(* IEC 61131-3 sources: daoli-st-library/_quarantine/R79, 13 files *)

(* ---- FC_DL_CalIsLeapYear.st ---- *)
(*==============================================================================
 * 组件名称 : FC_DL_CalIsLeapYear ｜ 子库 : DL_MathData ｜ v1.0.0 ｜ 2026-11-24
 * 平台     : CODESYS 3.5 / TwinCAT 3 / InoProShop / Machine Expert（纯 IEC，无厂商库）
 * 功能简介 : 公历（格里高利历）闰年判定 —— 能被 4 整除且不能被 100 整除，或能被 400
 *            整除即为闰年。纯整数取余，无浮点、无日历库依赖。
 * 契约     : 返回 TRUE=闰年；nYear < 1583（格里高利历起点）返回 FALSE 且
 *            bValid := FALSE —— 儒略历闰年口径与本件不同，域外一律不认。
 *            纯函数无状态，同输入同输出。
 * 依赖     : 无 DL_ 内部依赖（R16 自足实现），无标准库函数调用
 * 错误码   : R297 零码位范式：eErr 恒 0，仅以 bError / bValid 表达（本件结构性不置 bError）
 * 红线自检 : R1 零全局 R2 零%I/%Q R3 纯IEC R4 取余无除法歧义、域闸先判年份
 *            R5 双语注释 R6 N/A（无状态机）R7 N/A（无定时器/沿实例）
 *            R10 无类型转换 R11 全声明行分号 R15 标识符零保留字冲突 R18 N/A（无 bReset）
 * 修订历史 : 2026-11-24 R79-A 首版（日历算术族 1/9）
 *============================================================================*)
FUNCTION FC_DL_CalIsLeapYear : BOOL
VAR_INPUT
    nYear    : DINT;    // 待判定公历年，有效域 1583 及以上 [年] / Gregorian year to test, valid from 1583 [year]
END_VAR
VAR_OUTPUT
    eErr     : UDINT;   // 错误码，零码位范式恒 0 / error id, always zero under the zero-code rule
    bError   : BOOL;    // 故障标志，本件结构性不置位 / fault flag, never raised by this component
    bValid   : BOOL;    // 年份落在格里高利历域内为真 / TRUE when the year is inside the Gregorian domain
END_VAR
VAR CONSTANT
    DL_GREG_START : DINT := 1583;   // 格里高利历起点年 [年] / first Gregorian year [year]
    DL_STEP4      : DINT := 4;      // 闰年基本步长 [年] / base leap step [year]
    DL_STEP100    : DINT := 100;    // 世纪基数 [年] / century radix [year]
    DL_STEP400    : DINT := 400;    // 四世纪基数 [年] / four century radix [year]
    DL_ZERO       : DINT := 0;      // 整数零哨兵 [无量纲] / integer zero sentinel [dimensionless]
END_VAR
VAR
    nMod4    : DINT;    // 年份除 4 的余数 [无量纲] / remainder of the year divided by four [dimensionless]
    nMod100  : DINT;    // 年份除 100 的余数 [无量纲] / remainder of the year divided by one hundred [dimensionless]
    nMod400  : DINT;    // 年份除 400 的余数 [无量纲] / remainder of the year divided by four hundred [dimensionless]
END_VAR

// 段 1｜出口预置：任何路径下结果确定 / segment 1, preset the exit so that every path is deterministic
FC_DL_CalIsLeapYear := FALSE;   // 缺省非闰年 / default is not a leap year
eErr   := 0;                    // 零码位范式 / zero-code rule
bError := FALSE;                // 本件不产生故障级 / this component raises no fault
bValid := FALSE;                // 域闸通过前不认结果 / the result stays unusable until the domain gate passes

// 段 2｜域闸：1583 之前属儒略历，闰年口径不同，直接拒绝 / segment 2, the domain gate rejects years before 1583
IF nYear < DL_GREG_START THEN
    RETURN;                     // 返回 FALSE 且 bValid 保持 FALSE / return FALSE with bValid still FALSE
END_IF
bValid := TRUE;                 // 年份入域，结果可用 / the year is inside the domain, the result is usable

// 段 3｜闰年判据：先取三个余数，再做布尔合成（避免重复取余） / segment 3, the leap rule on three remainders
nMod4   := nYear MOD DL_STEP4;      // 4 年周期余数 / remainder against four years
nMod100 := nYear MOD DL_STEP100;    // 100 年周期余数 / remainder against one hundred years
nMod400 := nYear MOD DL_STEP400;    // 400 年周期余数 / remainder against four hundred years
IF ((nMod4 = DL_ZERO) AND (nMod100 <> DL_ZERO)) OR (nMod400 = DL_ZERO) THEN
    FC_DL_CalIsLeapYear := TRUE;    // 整除 4 且不整除 100，或整除 400 / divisible by four but not by one hundred, or divisible by four hundred
END_IF
END_FUNCTION

(* ---- FC_DL_CalIsoWeekNo.st ---- *)
(*==============================================================================
 * 组件名称 : FC_DL_CalIsoWeekNo ｜ 子库 : DL_MathData ｜ v1.0.0 ｜ 2026-11-24
 * 平台     : CODESYS 3.5 / TwinCAT 3 / InoProShop / Machine Expert（纯 IEC，无厂商库）
 * 功能简介 : ISO 8601 周号 —— 周一起算，含 1 月 4 日的那一周为第 1 周。核心式
 *            week = (年内序号 − ISO 星期 + 10) DIV 7。跨年归属单独处理：算出 0 即属
 *            上年末周，算出超过当年周数即属次年 W1，并用出参 nWeekYear 标明归属年。
 * 契约     : 返回周号 1~53，nWeekYear 为归属年；nYear < 1583、月份或日越界时返回 -1、
 *            bError := TRUE、nWeekYear := 0。纯函数无状态。
 * 依赖     : 无 DL_ 内部依赖（R16 自足实现），无标准库函数调用
 * 错误码   : R297 零码位范式：eErr 恒 0，仅以 bError / bValid 表达
 * 红线自检 : R1 零全局 R2 零%I/%Q R3 纯IEC R4 三层域闸、取余操作数恒非负、除数为常量 7
 *            R5 双语注释 R6 N/A（无状态机）R7 N/A（无定时器/沿实例）
 *            R10 无类型转换 R11 全声明行分号 R15 标识符零保留字冲突 R18 N/A（无 bReset）
 * 遗留假设 : 53 周年判据按 ISO 官方口径取「1 月 1 日为周四」或「闰年且 1 月 1 日为周三」；
 *            该两式与「12 月 31 日落在第 53 周」等价，本件用前者以便直接复用 1 月 1 日序数。
 * 修订历史 : 2026-11-24 R79-A 首版（日历算术族 6/9）
 *============================================================================*)
FUNCTION FC_DL_CalIsoWeekNo : DINT
VAR_INPUT
    nYear      : DINT;  // 公历年，域闸 1583 及以上 [年] / Gregorian year, domain starts at 1583 [year]
    nMonth     : DINT;  // 月份 1~12 [月] / month from one to twelve [month]
    nDay       : DINT;  // 日 1~当月天数 [天] / day from one to the month length [day]
END_VAR
VAR_OUTPUT
    eErr       : UDINT; // 错误码，零码位范式恒 0 / error id, always zero under the zero-code rule
    bError     : BOOL;  // 日期非法或域外为真 / TRUE when the date is illegal or out of domain
    bValid     : BOOL;  // 结果可用标志 / result usable flag
    nWeekYear  : DINT;  // 周号归属年，故障时 0 [年] / year owning the ISO week, zero on fault [year]
END_VAR
VAR CONSTANT
    DL_GREG_START : DINT := 1583;   // 格里高利历起点年 [年] / first Gregorian year [year]
    DL_MONTH_MIN  : DINT := 1;      // 月份与日的下界 [月] / lower bound of the month and the day [month]
    DL_MONTH_MAX  : DINT := 12;     // 月份上界 [月] / upper month bound [month]
    DL_DAYS_COMMON : DINT := 365;   // 平年天数 [天] / days in a common year [day]
    DL_DAYS_FEB   : DINT := 28;     // 平年 2 月天数 [天] / February days in a common year [day]
    DL_DAYS_30    : DINT := 30;     // 小月天数 [天] / days in a short month [day]
    DL_DAYS_31    : DINT := 31;     // 大月天数 [天] / days in a long month [day]
    DL_STEP4      : DINT := 4;      // 闰年基本步长 [年] / base leap step [year]
    DL_STEP100    : DINT := 100;    // 世纪基数 [年] / century radix [year]
    DL_STEP400    : DINT := 400;    // 四世纪基数 [年] / four century radix [year]
    DL_WEEK_MOD   : DINT := 7;      // 星期与周号的基数 [天] / weekday and week radix [day]
    DL_WEEK_MIN   : DINT := 1;      // 周号下界 [周] / lower bound of the week number [week]
    DL_WEEK_BASE  : DINT := 52;     // 每年基础周数，53 周为特例 [周] / base weeks per year, fifty three is the exception [week]
    DL_WEEK_OFF   : DINT := 10;     // 周号式的固定偏移 [天] / fixed offset of the week formula [day]
    DL_JAN1_DOW53A : DINT := 4;     // 1 月 1 日周四 → 53 周 [星期序号] / Thursday first of January gives fifty three weeks
    DL_JAN1_DOW53B : DINT := 3;     // 闰年 1 月 1 日周三 → 53 周 [星期序号] / Wednesday first of January in a leap year gives fifty three weeks
    DL_ZERO       : DINT := 0;      // 整数零哨兵 [无量纲] / integer zero sentinel [dimensionless]
END_VAR
VAR
    bLeap      : BOOL;  // 当年是否闰年 / whether the year is a leap year
    bLeapPrev  : BOOL;  // 上一年是否闰年 / whether the previous year is a leap year
    nDaysInMon : DINT;  // 当月实际天数 [天] / actual length of the month [day]
    nDaysYear  : DINT;  // 当年总天数 365 或 366 [天] / total days of the year [day]
    nDaysPrev  : DINT;  // 上年总天数 365 或 366 [天] / total days of the previous year [day]
    nA         : DINT;  // 月份压缩偏置 0 或 1 / month compression offset, zero or one
    nY2        : DINT;  // 儒略式内的世纪内年份 / shifted year inside the Julian formula
    nM2        : DINT;  // 儒略式内的三月基月份 / March based month inside the Julian formula
    nJdn       : DINT;  // 目标日期的儒略日序数 [日] / Julian day number of the requested date [day]
    nJdnJan1   : DINT;  // 同年 1 月 1 日的儒略日序数 [日] / Julian day number of January the first [day]
    nDowJan1   : DINT;  // 1 月 1 日的 ISO 星期 1~7 [星期序号] / ISO weekday of January the first, one to seven
    nW         : DINT;  // 目标日期的 ISO 星期 1~7 [星期序号] / ISO weekday of the requested date, one to seven
    nOrd       : DINT;  // 年内序号 1~366 [天] / day of year, one to three hundred sixty six [day]
    nWeek      : DINT;  // 周号中间量 0~54 [周] / week interim value, zero to fifty four [week]
    nWeeksYear : DINT;  // 当年 ISO 周数 52 或 53 [周] / ISO weeks in the year, fifty two or fifty three [week]
END_VAR

// 段 1｜出口预置 / segment 1, preset the exit
FC_DL_CalIsoWeekNo := -1;       // 缺省无效哨兵 / default invalid sentinel
eErr       := 0;                // 零码位范式 / zero-code rule
bError     := FALSE;            // 预置无故障 / preset no fault
bValid     := FALSE;            // 域闸前不认结果 / unusable until the domain gates pass
nWeekYear  := 0;                // 归属年清零 / clear the owning year

// 段 2｜域闸：年份 → 月份 → 日（含闰年 2 月） / segment 2, the three domain gates
bLeap := (((nYear MOD DL_STEP4) = DL_ZERO) AND ((nYear MOD DL_STEP100) <> DL_ZERO)) OR ((nYear MOD DL_STEP400) = DL_ZERO);
nDaysYear := DL_DAYS_COMMON;
IF bLeap THEN
    nDaysYear := DL_DAYS_COMMON + 1;    // 闰年多一天 / a leap year carries one extra day
END_IF
IF (nYear < DL_GREG_START) OR (nMonth < DL_MONTH_MIN) OR (nMonth > DL_MONTH_MAX) THEN
    bError := TRUE;             // 年份或月份越界 / the year or the month is out of range
    RETURN;
END_IF
IF nMonth = 2 THEN
    nDaysInMon := DL_DAYS_FEB;          // 平年 2 月 / common February
    IF bLeap THEN
        nDaysInMon := DL_DAYS_FEB + 1;  // 闰年 2 月 / leap February
    END_IF
ELSIF (nMonth = 4) OR (nMonth = 6) OR (nMonth = 9) OR (nMonth = 11) THEN
    nDaysInMon := DL_DAYS_30;           // 小月 / short month
ELSE
    nDaysInMon := DL_DAYS_31;           // 大月 / long month
END_IF
IF (nDay < DL_MONTH_MIN) OR (nDay > nDaysInMon) THEN
    bError := TRUE;             // 日超出当月天数 / the day exceeds the month length
    RETURN;
END_IF

// 段 3｜两个儒略日序数：目标日期与同年 1 月 1 日 / segment 3, two Julian day numbers
nA   := (14 - nMonth) / 12;                                  // 1、2 月折入上一年 / January and February fold backwards
nY2  := nYear + 4800 - nA;                                   // 世纪内年份偏置 / shifted year
nM2  := nMonth + 12 * nA - 3;                                // 三月基月份 / March based month
nJdn := nDay + (153 * nM2 + 2) / 5 + 365 * nY2 + nY2 / DL_STEP4 - nY2 / DL_STEP100 + nY2 / DL_STEP400 - 32045;
nJdnJan1 := 307 + 365 * (nYear + 4799) + (nYear + 4799) / DL_STEP4 - (nYear + 4799) / DL_STEP100 + (nYear + 4799) / DL_STEP400 - 32045;
nOrd := nJdn - nJdnJan1 + 1;                                 // 年内序号 / day of year
nW   := (nJdn MOD DL_WEEK_MOD) + 1;                           // ISO 星期 1=周一 … 7=周日 / ISO weekday

// 段 4｜周号主式与当年周数：53 周须 1 月 1 日为周四，或闰年且为周三 / segment 4, the week formula and the year length
nWeek := (nOrd - nW + DL_WEEK_OFF) / DL_WEEK_MOD;             // 0~54 中间值 / interim value
nDowJan1 := (nJdnJan1 MOD DL_WEEK_MOD) + 1;                   // 1 月 1 日的 ISO 星期 / ISO weekday of January the first
nWeeksYear := DL_WEEK_BASE;                                   // 缺省 52 周 / default fifty two weeks
IF (nDowJan1 = DL_JAN1_DOW53A) OR (bLeap AND (nDowJan1 = DL_JAN1_DOW53B)) THEN
    nWeeksYear := DL_WEEK_BASE + 1;                           // 该年为 53 周 / the year carries fifty three weeks
END_IF

// 段 5｜跨年归属：0 归上年末周，超年周数归次年 W1 / segment 5, the two cross year branches
nWeekYear := nYear;
IF nWeek < DL_WEEK_MIN THEN
    bLeapPrev := ((((nYear - 1) MOD DL_STEP4) = DL_ZERO) AND (((nYear - 1) MOD DL_STEP100) <> DL_ZERO)) OR (((nYear - 1) MOD DL_STEP400) = DL_ZERO);
    nDaysPrev := DL_DAYS_COMMON;
    IF bLeapPrev THEN
        nDaysPrev := DL_DAYS_COMMON + 1;    // 上年为闰年 / the previous year is a leap year
    END_IF
    nWeek     := (nOrd + nDaysPrev - nW + DL_WEEK_OFF) / DL_WEEK_MOD;   // 换算到上年的序数 / rebase onto the previous year
    nWeekYear := nYear - 1;                                             // 归属上年 / owned by the previous year
ELSIF nWeek > nWeeksYear THEN
    nWeek     := (nOrd - nDaysYear - nW + DL_WEEK_OFF) / DL_WEEK_MOD;   // 换算到次年的序数 / rebase onto the next year
    IF nWeek < DL_WEEK_MIN THEN
        nWeek := DL_WEEK_MIN;                                          // 结构性必为 1，兜底防御 / always one, kept as a guard
    END_IF
    nWeekYear := nYear + 1;                                             // 归属次年 / owned by the next year
END_IF

// 段 6｜出口 / segment 6, exit
FC_DL_CalIsoWeekNo := nWeek;    // 1~53 / one to fifty three
bValid := TRUE;                 // 结果可用 / the result is usable
END_FUNCTION

(* ---- FC_DL_CalMonthDays.st ---- *)
(*==============================================================================
 * 组件名称 : FC_DL_CalMonthDays ｜ 子库 : DL_MathData ｜ v1.0.0 ｜ 2026-11-24
 * 平台     : CODESYS 3.5 / TwinCAT 3 / InoProShop / Machine Expert（纯 IEC，无厂商库）
 * 功能简介 : 给定公历年月，返回该月天数；2 月按闰年判据取 28 或 29，其余月固定 30/31。
 *            纯整数实现，闰年判据内联自足，不调用同族其他件。
 * 契约     : 返回 1~31 为合法天数；nMonth 越界（<1 或 >12）返回 0 且 bError := TRUE。
 *            nYear < 1583 时 2 月按非闰年（28）计数 —— 儒略历口径不入本件，见遗留假设。
 * 依赖     : 无 DL_ 内部依赖（R16 自足实现），无标准库函数调用
 * 错误码   : R297 零码位范式：eErr 恒 0，仅以 bError / bValid 表达
 * 红线自检 : R1 零全局 R2 零%I/%Q R3 纯IEC R4 月份域闸先行、取余无除零面
 *            R5 双语注释 R6 N/A（无状态机）R7 N/A（无定时器/沿实例）
 *            R10 无类型转换 R11 全声明行分号 R15 标识符零保留字冲突 R18 N/A（无 bReset）
 * 遗留假设 : 格里高利历起点之前的 2 月按 28 天计；该域需 29 天的场合请先自查历法归属。
 * 修订历史 : 2026-11-24 R79-A 首版（日历算术族 2/9）
 *============================================================================*)
FUNCTION FC_DL_CalMonthDays : DINT
VAR_INPUT
    nYear     : DINT;   // 公历年，仅供 2 月闰年判定 [年] / Gregorian year used by the February leap test [year]
    nMonth    : DINT;   // 月份 1~12，越界即故障 [月] / month from one to twelve, out of range is a fault [month]
END_VAR
VAR_OUTPUT
    eErr      : UDINT;  // 错误码，零码位范式恒 0 / error id, always zero under the zero-code rule
    bError    : BOOL;   // 月份越界为真，返回 0 / TRUE when the month is out of range, the result is zero
    bValid    : BOOL;   // 结果可用标志 / result usable flag
END_VAR
VAR CONSTANT
    DL_MONTH_MIN  : DINT := 1;      // 月份下界 [月] / lower month bound [month]
    DL_MONTH_MAX  : DINT := 12;     // 月份上界 [月] / upper month bound [month]
    DL_DAYS_31    : DINT := 31;     // 大月天数 [天] / days in a long month [day]
    DL_DAYS_30    : DINT := 30;     // 小月天数 [天] / days in a short month [day]
    DL_DAYS_FEB   : DINT := 28;     // 平年 2 月天数 [天] / February days in a common year [day]
    DL_GREG_START : DINT := 1583;   // 格里高利历起点年 [年] / first Gregorian year [year]
    DL_STEP4      : DINT := 4;      // 闰年基本步长 [年] / base leap step [year]
    DL_STEP100    : DINT := 100;    // 世纪基数 [年] / century radix [year]
    DL_STEP400    : DINT := 400;    // 四世纪基数 [年] / four century radix [year]
    DL_ZERO       : DINT := 0;      // 整数零哨兵 [无量纲] / integer zero sentinel [dimensionless]
END_VAR
VAR
    bLeap     : BOOL;   // 当年是否闰年 / whether the year is a leap year
END_VAR

// 段 1｜出口预置 / segment 1, preset the exit
FC_DL_CalMonthDays := 0;        // 缺省 0 天 / default zero days
eErr   := 0;                    // 零码位范式 / zero-code rule
bError := FALSE;                // 预置无故障 / preset no fault
bValid := FALSE;                // 域闸前不认结果 / unusable until the domain gate passes

// 段 2｜月份域闸：唯一故障出口 / segment 2, the month domain gate is the only fault exit
IF (nMonth < DL_MONTH_MIN) OR (nMonth > DL_MONTH_MAX) THEN
    bError := TRUE;             // 月份越界 / the month is out of range
    RETURN;                     // 返回 0 / return zero
END_IF
bValid := TRUE;                 // 月份入域 / the month is inside the domain

// 段 3｜闰年判据（内联自足，不跨件调用） / segment 3, the leap test implemented inline
bLeap := FALSE;
IF nYear >= DL_GREG_START THEN
    bLeap := (((nYear MOD DL_STEP4) = DL_ZERO) AND ((nYear MOD DL_STEP100) <> DL_ZERO)) OR ((nYear MOD DL_STEP400) = DL_ZERO);
END_IF

// 段 4｜月长选择：2 月单列，30 天月枚举，其余一律 31 天 / segment 4, month length selection
IF nMonth = 2 THEN
    IF bLeap THEN
        FC_DL_CalMonthDays := DL_DAYS_FEB + 1;     // 闰年 2 月 29 天 / twenty nine days in a leap February
    ELSE
        FC_DL_CalMonthDays := DL_DAYS_FEB;         // 平年 2 月 28 天 / twenty eight days otherwise
    END_IF
ELSIF (nMonth = 4) OR (nMonth = 6) OR (nMonth = 9) OR (nMonth = 11) THEN
    FC_DL_CalMonthDays := DL_DAYS_30;              // 4/6/9/11 月为 30 天 / thirty day months
ELSE
    FC_DL_CalMonthDays := DL_DAYS_31;              // 其余为 31 天 / the rest have thirty one days
END_IF
END_FUNCTION

(* ---- FC_DL_CalMonthEndDate.st ---- *)
(*==============================================================================
 * 组件名称 : FC_DL_CalMonthEndDate ｜ 子库 : DL_MathData ｜ v1.0.1 ｜ 2026-11-24
 * 平台     : CODESYS 3.5 / TwinCAT 3 / InoProShop / Machine Expert（纯 IEC，无厂商库）
 * 功能简介 : 给定公历年月，出参返回该月最后一天的日号（月末日期）。月度报表切日、
 *            月累计清零、月末结账触发都以本件为唯一口径。2 月按闰年判据取 28 / 29。
 * 契约     : 合法时返回 TRUE 并写出 nLastDay（1~31）；nMonth 越界或 nYear < 1583 时
 *            返回 FALSE、bError := TRUE、nLastDay := 0。纯函数无状态。
 * 依赖     : 无 DL_ 内部依赖（R16 自足实现），无标准库函数调用
 * 错误码   : R297 零码位范式：eErr 恒 0，仅以 bError / bValid 表达
 * 红线自检 : R1 零全局 R2 零%I/%Q R3 纯IEC R4 年份与月份双域闸、取余无除零面
 *            R5 双语注释 R6 N/A（无状态机）R7 N/A（无定时器/沿实例）
 *            R10 无类型转换 R11 全声明行分号 R15 标识符零保留字冲突 R18 N/A（无 bReset）
 * 修订历史 : 2026-11-24 R79-A 首版（日历算术族 9/9）
 *            2026-11-24  v1.0.1  R79/P4：补年份上界闸 DL_GREG_LAST=9999（原仅下界 1583）
 *============================================================================*)
FUNCTION FC_DL_CalMonthEndDate : BOOL
VAR_INPUT
    nYear     : DINT;   // 公历年，域闸 1583 及以上 [年] / Gregorian year, domain starts at 1583 [year]
    nMonth    : DINT;   // 月份 1~12 [月] / month from one to twelve [month]
END_VAR
VAR_OUTPUT
    eErr      : UDINT;  // 错误码，零码位范式恒 0 / error id, always zero under the zero-code rule
    bError    : BOOL;   // 年份或月份越界为真 / TRUE when the year or the month is out of range
    bValid    : BOOL;   // 出参可用标志 / TRUE when the output is usable
    nLastDay  : DINT;   // 该月最后一天的日号 1~31，故障时 0 [天] / last day of the month, zero on fault [day]
END_VAR
VAR CONSTANT
    DL_GREG_START : DINT := 1583;   // 格里高利历起点年 [年] / first Gregorian year [year]
    DL_GREG_LAST  : DINT := 9999;   // 年份上界（v1.0.1 补：防 int64/日期串溢出）[年] / Upper year bound added in v1.0.1 [year]
    DL_MONTH_MIN  : DINT := 1;      // 月份下界 [月] / lower month bound [month]
    DL_MONTH_MAX  : DINT := 12;     // 月份上界 [月] / upper month bound [month]
    DL_DAYS_FEB   : DINT := 28;     // 平年 2 月天数 [天] / February days in a common year [day]
    DL_DAYS_30    : DINT := 30;     // 小月天数 [天] / days in a short month [day]
    DL_DAYS_31    : DINT := 31;     // 大月天数 [天] / days in a long month [day]
    DL_STEP4      : DINT := 4;      // 闰年基本步长 [年] / base leap step [year]
    DL_STEP100    : DINT := 100;    // 世纪基数 [年] / century radix [year]
    DL_STEP400    : DINT := 400;    // 四世纪基数 [年] / four century radix [year]
    DL_ZERO       : DINT := 0;      // 整数零哨兵 [无量纲] / integer zero sentinel [dimensionless]
END_VAR
VAR
    bLeap     : BOOL;   // 当年是否闰年 / whether the year is a leap year
END_VAR

// 段 1｜出口预置 / segment 1, preset the exit
FC_DL_CalMonthEndDate := FALSE;     // 缺省失败 / default failure
eErr      := 0;                     // 零码位范式 / zero-code rule
bError    := FALSE;                 // 预置无故障 / preset no fault
bValid    := FALSE;                 // 域闸前不认出参 / the output is unusable until the gates pass
nLastDay  := 0;                     // 日号清零 / clear the day number

// 段 2｜域闸：年份 → 月份 / segment 2, the year and the month gates
IF ((nYear < DL_GREG_START) OR (nYear > DL_GREG_LAST)) OR (nMonth < DL_MONTH_MIN) OR (nMonth > DL_MONTH_MAX) THEN
    bError := TRUE;                 // 年份或月份越界 / the year or the month is out of range
    RETURN;                         // 出参保持 0 / the output stays zero
END_IF

// 段 3｜闰年判据（内联自足） / segment 3, the leap test implemented inline
bLeap := (((nYear MOD DL_STEP4) = DL_ZERO) AND ((nYear MOD DL_STEP100) <> DL_ZERO)) OR ((nYear MOD DL_STEP400) = DL_ZERO);

// 段 4｜月末日号：2 月单列，30 天月枚举，其余 31 天 / segment 4, the last day selection
IF nMonth = 2 THEN
    nLastDay := DL_DAYS_FEB;        // 平年 2 月 / common February
    IF bLeap THEN
        nLastDay := DL_DAYS_FEB + 1;    // 闰年 2 月 / leap February
    END_IF
ELSIF (nMonth = 4) OR (nMonth = 6) OR (nMonth = 9) OR (nMonth = 11) THEN
    nLastDay := DL_DAYS_30;         // 小月 / short month
ELSE
    nLastDay := DL_DAYS_31;         // 大月 / long month
END_IF

// 段 5｜出口 / segment 5, exit
bValid := TRUE;                     // 出参可用 / the output is usable
FC_DL_CalMonthEndDate := TRUE;      // 求解成功 / the request succeeded
END_FUNCTION

(* ---- FC_DL_CalWeekdayIndex.st ---- *)
(*==============================================================================
 * 组件名称 : FC_DL_CalWeekdayIndex ｜ 子库 : DL_MathData ｜ v1.0.0 ｜ 2026-11-24
 * 平台     : CODESYS 3.5 / TwinCAT 3 / InoProShop / Machine Expert（纯 IEC，无厂商库）
 * 功能简介 : 公历日期的 ISO 星期序号 —— 0=周一 … 6=周日。用儒略日序数取余实现：
 *            JDN MOD 7 恰为「周一为 0」的序号（JDN 0 落在周一），纯整数、无浮点。
 * 契约     : 返回 0~6；nYear < 1583、nMonth 不在 1~12、nDay 超出当月天数时返回 -1 且
 *            bError := TRUE。纯函数无状态，同输入同输出。
 * 依赖     : 无 DL_ 内部依赖（R16 自足实现），无标准库函数调用
 * 错误码   : R297 零码位范式：eErr 恒 0，仅以 bError / bValid 表达
 * 红线自检 : R1 零全局 R2 零%I/%Q R3 纯IEC R4 三层域闸先行、取余操作数恒非负
 *            R5 双语注释 R6 N/A（无状态机）R7 N/A（无定时器/沿实例）
 *            R10 无类型转换 R11 全声明行分号 R15 标识符零保留字冲突 R18 N/A（无 bReset）
 * 遗留假设 : 1583 年以前走儒略历，儒略日序数与格里高利历存在跳日差，故设域闸下限。
 * 修订历史 : 2026-11-24 R79-A 首版（日历算术族 5/9）
 *============================================================================*)
FUNCTION FC_DL_CalWeekdayIndex : DINT
VAR_INPUT
    nYear     : DINT;   // 公历年，域闸 1583 及以上 [年] / Gregorian year, domain starts at 1583 [year]
    nMonth    : DINT;   // 月份 1~12 [月] / month from one to twelve [month]
    nDay      : DINT;   // 日 1~当月天数 [天] / day from one to the month length [day]
END_VAR
VAR_OUTPUT
    eErr      : UDINT;  // 错误码，零码位范式恒 0 / error id, always zero under the zero-code rule
    bError    : BOOL;   // 日期不存在或域外为真 / TRUE when the date is invalid or out of domain
    bValid    : BOOL;   // 结果可用标志 / result usable flag
END_VAR
VAR CONSTANT
    DL_GREG_START : DINT := 1583;   // 格里高利历起点年 [年] / first Gregorian year [year]
    DL_MONTH_MIN  : DINT := 1;      // 月份与日的下界 [月] / lower bound of the month and the day [month]
    DL_MONTH_MAX  : DINT := 12;     // 月份上界 [月] / upper month bound [month]
    DL_DAYS_FEB   : DINT := 28;     // 平年 2 月天数 [天] / February days in a common year [day]
    DL_DAYS_30    : DINT := 30;     // 小月天数 [天] / days in a short month [day]
    DL_DAYS_31    : DINT := 31;     // 大月天数 [天] / days in a long month [day]
    DL_STEP4      : DINT := 4;      // 闰年基本步长 [年] / base leap step [year]
    DL_STEP100    : DINT := 100;    // 世纪基数 [年] / century radix [year]
    DL_STEP400    : DINT := 400;    // 四世纪基数 [年] / four century radix [year]
    DL_WEEK_MOD   : DINT := 7;      // 星期基数 [天] / weekday radix [day]
    DL_ZERO       : DINT := 0;      // 整数零哨兵 [无量纲] / integer zero sentinel [dimensionless]
END_VAR
VAR
    bLeap      : BOOL;  // 当年是否闰年 / whether the year is a leap year
    nDaysInMon : DINT;  // 当月实际天数 [天] / actual length of the month [day]
    nA         : DINT;  // 月份压缩偏置 0 或 1 / month compression offset, zero or one
    nY2        : DINT;  // 儒略式内的世纪内年份 / shifted year inside the Julian formula
    nM2        : DINT;  // 儒略式内的三月基月份 / March based month inside the Julian formula
    nJdn       : DINT;  // 目标日期的儒略日序数 [日] / Julian day number of the requested date [day]
END_VAR

// 段 1｜出口预置：缺省 -1 表示无效 / segment 1, preset the exit to minus one
FC_DL_CalWeekdayIndex := -1;    // 无效哨兵 / invalid sentinel
eErr   := 0;                    // 零码位范式 / zero-code rule
bError := FALSE;                // 预置无故障 / preset no fault
bValid := FALSE;                // 域闸前不认结果 / unusable until the domain gates pass

// 段 2｜域闸：年份 → 月份 → 日 / segment 2, three domain gates in sequence
IF (nYear < DL_GREG_START) OR (nMonth < DL_MONTH_MIN) OR (nMonth > DL_MONTH_MAX) THEN
    bError := TRUE;             // 年份或月份越界 / the year or the month is out of range
    RETURN;                     // 返回 -1 / return minus one
END_IF
bLeap := (((nYear MOD DL_STEP4) = DL_ZERO) AND ((nYear MOD DL_STEP100) <> DL_ZERO)) OR ((nYear MOD DL_STEP400) = DL_ZERO);
IF nMonth = 2 THEN
    nDaysInMon := DL_DAYS_FEB;          // 平年 2 月 / common February
    IF bLeap THEN
        nDaysInMon := DL_DAYS_FEB + 1;  // 闰年 2 月 / leap February
    END_IF
ELSIF (nMonth = 4) OR (nMonth = 6) OR (nMonth = 9) OR (nMonth = 11) THEN
    nDaysInMon := DL_DAYS_30;           // 小月 / short month
ELSE
    nDaysInMon := DL_DAYS_31;           // 大月 / long month
END_IF
IF (nDay < DL_MONTH_MIN) OR (nDay > nDaysInMon) THEN
    bError := TRUE;             // 日超出当月天数 / the day exceeds the month length
    RETURN;                     // 返回 -1 / return minus one
END_IF

// 段 3｜儒略日序数 / segment 3, the Julian day number
nA   := (14 - nMonth) / 12;                                  // 1、2 月折入上一年 / January and February fold backwards
nY2  := nYear + 4800 - nA;                                   // 世纪内年份偏置 / shifted year
nM2  := nMonth + 12 * nA - 3;                                // 三月基月份 / March based month
nJdn := nDay + (153 * nM2 + 2) / 5 + 365 * nY2 + nY2 / DL_STEP4 - nY2 / DL_STEP100 + nY2 / DL_STEP400 - 32045;

// 段 4｜出口：JDN 模 7 即「周一为 0」的 ISO 序号 / segment 4, JDN modulo seven is the Monday based index
FC_DL_CalWeekdayIndex := nJdn MOD DL_WEEK_MOD;   // 0=周一 … 6=周日 / zero equals Monday and six equals Sunday
bValid := TRUE;                                  // 日期合法，结果可用 / the date is legal and the result is usable
END_FUNCTION

(* ---- FC_DL_ChkSum8.st ---- *)
(*==============================================================================
 * 组件名称 : FC_DL_ChkSum8 ｜ 子库 : DL_Algo ｜ v1.0.0 ｜ 2026-11-24
 * 平台     : CODESYS 3.5 / TwinCAT 3 / InoProShop / Machine Expert（纯 IEC，无厂商库）
 * 功能简介 : 字节和校验（Sum-8 / LRC 的加和型）。全部字节求和后取模 256，返回单字节。
 *            仪表与老式 PLC 的 ASCII 协议最常用的帧尾校验之一。
 * 契约     : 返回 sum MOD 256；nLen 越界钳到 0~16；nLen = 0 返回 0。
 *            数组定长 ARRAY[1..16] OF BYTE（R17）。
 * 依赖     : 无 DL_ 内部依赖（R16 自足实现）；Standard.library: BYTE_TO_UDINT / UDINT_TO_BYTE
 * 错误码   : R297 零码位范式：eErr 恒 0，本件结构性不置 bError
 * 红线自检 : R1 零全局 R2 零%I/%Q R3 纯IEC R4 累加在 UDINT 域（16×255 远小于 2^32）、
 *            取模后再收窄到 BYTE，收窄前值必 < 256 ｜ R5 双语注释 R6 N/A（无状态机）
 *            R7 N/A（无定时器/沿实例）R10 标准转换 R11 全声明行分号
 *            R15 标识符零保留字冲突 R17 定长数组 R18 N/A（无 bReset）
 * 遗留假设 : 取模口径为 256（2 的幂），与 255 口径的 Fletcher 不同，对接协议前须核对。
 * 修订历史 : 2026-11-24 R79-A 首版（校验和族 4/8）
 *============================================================================*)
FUNCTION FC_DL_ChkSum8 : BYTE
VAR_INPUT
    aData   : ARRAY[1..16] OF BYTE;     // 待校验字节块，1..16 定长 [字节] / byte block of fixed length [byte]
    nLen    : INT;                      // 有效字节数 0~16，越界钳位 [字节] / effective length from zero to sixteen, clamped [byte]
END_VAR
VAR_OUTPUT
    eErr    : UDINT;                    // 错误码，零码位范式恒 0 / error id, always zero under the zero-code rule
    bError  : BOOL;                     // 故障标志，本件结构性不置位 / fault flag, never raised by this component
    bValid  : BOOL;                     // 结果可用标志，空块亦可用 / TRUE even for an empty block
END_VAR
VAR CONSTANT
    DL_LEN_MAX : INT := 16;             // 字节块定长上限 [字节] / fixed block capacity [byte]
    DL_LEN_MIN : INT := 0;              // 长度下界，0 合法 [字节] / lower length bound, zero is legal [byte]
    DL_ONE     : INT := 1;              // 数组首下标 [字节] / first array index [byte]
    DL_MOD256  : UDINT := 256;          // 取模基数 [无量纲] / the modulus
    DL_ZERO_U  : UDINT := 0;            // 无符号零哨兵 / unsigned zero sentinel
END_VAR
VAR
    nSum    : UDINT;                    // 宽域累加和，收窄前必 < 256 / wide accumulator, below 256 before narrowing
    nUse    : INT;                      // 钳位后的有效长度 [字节] / effective length after clamping [byte]
    i       : INT;                      // 遍历游标 [字节] / loop cursor [byte]
END_VAR

// 段 1｜出口预置 / segment 1, preset the exit
FC_DL_ChkSum8 := 16#00;             // 缺省 0 / default zero
eErr   := 0;                        // 零码位范式 / zero-code rule
bError := FALSE;                    // 本件不产生故障级 / this component raises no fault
bValid := TRUE;                     // 空块亦有定义 / an empty block is well defined
nSum   := DL_ZERO_U;                // 累加器清零 / clear the accumulator

// 段 2｜长度钳位：越界静默整形 / segment 2, clamp the length
nUse := nLen;
IF nUse < DL_LEN_MIN THEN
    nUse := DL_LEN_MIN;             // 下越界钳到 0 / clamp to zero
ELSIF nUse > DL_LEN_MAX THEN
    nUse := DL_LEN_MAX;             // 上越界钳到定长 / clamp to the fixed capacity
END_IF

// 段 3｜逐字节累加：16 个字节最大 4080，远小于 UDINT 上界 / segment 3, byte wise accumulation
FOR i := DL_ONE TO nUse DO
    nSum := nSum + BYTE_TO_UDINT(aData[i]);     // 宽域累加 / widen and accumulate
END_FOR

// 段 4｜出口：先取模再收窄，收窄时值必 < 256 / segment 4, take the modulus before narrowing
FC_DL_ChkSum8 := UDINT_TO_BYTE(nSum MOD DL_MOD256);
END_FUNCTION

(* ---- FC_DL_ChkXor8.st ---- *)
(*==============================================================================
 * 组件名称 : FC_DL_ChkXor8 ｜ 子库 : DL_Algo ｜ v1.0.0 ｜ 2026-11-24
 * 平台     : CODESYS 3.5 / TwinCAT 3 / InoProShop / Machine Expert（纯 IEC，无厂商库）
 * 功能简介 : 字节块异或校验（BCC / XOR-8）。全字节逐位异或，返回单字节结果。
 *            最简单的一类校验：对单比特翻转敏感，对字节顺序不敏感，
 *            常用于仪表 ASCII 协议的帧尾校验（模数恒为 256，天然无溢出）。
 * 契约     : 返回全字节异或值；nLen 越界钳到 0~16；nLen = 0 返回 0（空块异或为 0）。
 *            数组定长 ARRAY[1..16] OF BYTE（R17）。
 * 依赖     : 无 DL_ 内部依赖（R16 自足实现），无标准库函数调用
 * 错误码   : R297 零码位范式：eErr 恒 0，本件结构性不置 bError
 * 红线自检 : R1 零全局 R2 零%I/%Q R3 纯IEC R4 BYTE 异或天然模 256，无溢出面、
 *            长度先钳位后进循环 ｜ R5 双语注释 R6 N/A（无状态机）
 *            R7 N/A（无定时器/沿实例）R10 无类型转换 R11 全声明行分号
 *            R15 标识符零保留字冲突 R17 定长数组 R18 N/A（无 bReset）
 * 修订历史 : 2026-11-24 R79-A 首版（校验和族 3/8）
 *============================================================================*)
FUNCTION FC_DL_ChkXor8 : BYTE
VAR_INPUT
    aData   : ARRAY[1..16] OF BYTE;     // 待校验字节块，1..16 定长 [字节] / byte block of fixed length [byte]
    nLen    : INT;                      // 有效字节数 0~16，越界钳位 [字节] / effective length from zero to sixteen, clamped [byte]
END_VAR
VAR_OUTPUT
    eErr    : UDINT;                    // 错误码，零码位范式恒 0 / error id, always zero under the zero-code rule
    bError  : BOOL;                     // 故障标志，本件结构性不置位 / fault flag, never raised by this component
    bValid  : BOOL;                     // 结果可用标志，空块亦可用 / TRUE even for an empty block
END_VAR
VAR CONSTANT
    DL_LEN_MAX : INT := 16;             // 字节块定长上限 [字节] / fixed block capacity [byte]
    DL_LEN_MIN : INT := 0;              // 长度下界，0 合法 [字节] / lower length bound, zero is legal [byte]
    DL_ONE     : INT := 1;              // 数组首下标 [字节] / first array index [byte]
    DL_BYTE_ZERO : BYTE := 16#00;       // 字节零哨兵，异或单位元 / byte zero, the identity of the exclusive or
END_VAR
VAR
    nAcc    : BYTE;                     // 异或累加器 / exclusive or accumulator
    nUse    : INT;                      // 钳位后的有效长度 [字节] / effective length after clamping [byte]
    i       : INT;                      // 遍历游标 [字节] / loop cursor [byte]
END_VAR

// 段 1｜出口预置 / segment 1, preset the exit
FC_DL_ChkXor8 := DL_BYTE_ZERO;      // 缺省 0，空块异或即 0 / default zero, the identity of the operation
eErr   := 0;                        // 零码位范式 / zero-code rule
bError := FALSE;                    // 本件不产生故障级 / this component raises no fault
bValid := TRUE;                     // 空块亦有定义 / an empty block is well defined
nAcc   := DL_BYTE_ZERO;             // 累加器取异或单位元 / seed the accumulator with the identity

// 段 2｜长度钳位：越界静默整形 / segment 2, clamp the length
nUse := nLen;
IF nUse < DL_LEN_MIN THEN
    nUse := DL_LEN_MIN;             // 下越界钳到 0 / clamp to zero
ELSIF nUse > DL_LEN_MAX THEN
    nUse := DL_LEN_MAX;             // 上越界钳到定长 / clamp to the fixed capacity
END_IF

// 段 3｜逐字节异或：BYTE 域内运算，天然模 256 / segment 3, byte wise exclusive or
FOR i := DL_ONE TO nUse DO
    nAcc := nAcc XOR aData[i];      // 异或累积 / accumulate by exclusive or
END_FOR

// 段 4｜出口 / segment 4, exit
FC_DL_ChkXor8 := nAcc;              // 单字节结果 / the single byte result
END_FUNCTION

(* ---- FC_DL_GeoLineIntersectXY.st ---- *)
(*==============================================================================
 * 组件名称 : FC_DL_GeoLineIntersectXY ｜ 子库 : DL_MathData ｜ v1.0.0 ｜ 2026-11-24
 * 平台     : CODESYS 3.5 / TwinCAT 3 / InoProShop / Machine Expert（纯 IEC，无厂商库）
 * 功能简介 : 两线段求交点（参数式）。以行列式解出 t、u 两个线段参数，二者都落在 [0,1]
 *            才认为线段真实相交。用于视觉十字标定、激光对刀、两轴限位线交叉判定。
 * 契约     : 相交返回 TRUE 并写出 fX / fY；平行（|denom| < 1.0E-9）返回 FALSE 且
 *            bError := TRUE（几何病态）；共面但交点落在线段延长线上返回 FALSE 且
 *            bError := FALSE（正常无交点，不得当故障上报）。
 * 依赖     : 无 DL_ 内部依赖（R16 自足实现）；Standard.library: ABS
 * 错误码   : R297 零码位范式：eErr 恒 0，仅以 bError / bValid 表达
 * 红线自检 : R1 零全局 R2 零%I/%Q R3 纯IEC R4 除法前判 |denom| 容差、NaN 自反判据、
 *            无穷上界 ｜ R5 双语注释 R6 N/A（无状态机）R7 N/A（无定时器/沿实例）
 *            R10 无类型转换 R11 全声明行分号 R15 标识符零保留字冲突 R18 N/A（无 bReset）
 * 遗留假设 : 参数域容差取 1.0E-9，端点恰好落在对方端点上的情形判为相交（含边界）。
 * 修订历史 : 2026-11-24 R79-A 首版（平面几何族 2/8）
 *============================================================================*)
FUNCTION FC_DL_GeoLineIntersectXY : BOOL
VAR_INPUT
    fAx     : LREAL;    // 线段一 起点 X [mm] / start X of the first segment [mm]
    fAy     : LREAL;    // 线段一 起点 Y [mm] / start Y of the first segment [mm]
    fBx     : LREAL;    // 线段一 终点 X [mm] / end X of the first segment [mm]
    fBy     : LREAL;    // 线段一 终点 Y [mm] / end Y of the first segment [mm]
    fCx     : LREAL;    // 线段二 起点 X [mm] / start X of the second segment [mm]
    fCy     : LREAL;    // 线段二 起点 Y [mm] / start Y of the second segment [mm]
    fDx     : LREAL;    // 线段二 终点 X [mm] / end X of the second segment [mm]
    fDy     : LREAL;    // 线段二 终点 Y [mm] / end Y of the second segment [mm]
END_VAR
VAR_OUTPUT
    eErr    : UDINT;    // 错误码，零码位范式恒 0 / error id, always zero under the zero-code rule
    bError  : BOOL;     // 平行或非有限输入为真 / TRUE on parallel lines or non finite inputs
    bValid  : BOOL;     // 交点可用标志 / TRUE when the intersection point is usable
    fX      : LREAL;    // 交点 X 坐标，无交点时 0 [mm] / intersection X, zero when there is none [mm]
    fY      : LREAL;    // 交点 Y 坐标，无交点时 0 [mm] / intersection Y, zero when there is none [mm]
END_VAR
VAR CONSTANT
    DL_EPS      : LREAL := 1.0E-9;      // 行列式容差，小于它判为平行 [无量纲] / determinant tolerance, below it the lines are parallel
    DL_FIN_LIM  : LREAL := 1.0E308;     // 有限性上界 [无量纲] / finiteness ceiling
    DL_ONE      : LREAL := 1.0;         // 参数域上界 / upper bound of the segment parameter
    DL_ZERO_L   : LREAL := 0.0;         // 实数零哨兵 / real zero sentinel
END_VAR
VAR
    fD1x    : LREAL;    // 线段一方向 X 分量 B−A [mm] / direction X of the first segment [mm]
    fD1y    : LREAL;    // 线段一方向 Y 分量 B−A [mm] / direction Y of the first segment [mm]
    fD2x    : LREAL;    // 线段二方向 X 分量 D−C [mm] / direction X of the second segment [mm]
    fD2y    : LREAL;    // 线段二方向 Y 分量 D−C [mm] / direction Y of the second segment [mm]
    fDen    : LREAL;    // 两方向叉积（行列式）[mm²] / cross product of the two directions [mm²]
    fT      : LREAL;    // 线段一上的参数 [无量纲] / parameter along the first segment
    fU      : LREAL;    // 线段二上的参数 [无量纲] / parameter along the second segment
END_VAR

// 段 1｜出口预置 / segment 1, preset the exit
FC_DL_GeoLineIntersectXY := FALSE;  // 缺省无交点 / default no intersection
eErr   := 0;                        // 零码位范式 / zero-code rule
bError := FALSE;                    // 预置无故障 / preset no fault
bValid := FALSE;                    // 求解完成前不认交点 / the point is unusable until the solve ends
fX     := DL_ZERO_L;                // X 清零 / clear X
fY     := DL_ZERO_L;                // Y 清零 / clear Y

// 段 2｜非有限闸：八个坐标任一为 NaN 即拒 / segment 2, the non finite gate
IF (fAx <> fAx) OR (fAy <> fAy) OR (fBx <> fBx) OR (fBy <> fBy) OR (fCx <> fCx) OR (fCy <> fCy) OR (fDx <> fDx) OR (fDy <> fDy) THEN
    bError := TRUE;                 // 含非数输入 / a not a number input was seen
    RETURN;
END_IF

// 段 3｜方向与行列式：denom 为 0 即两线平行或重合 / segment 3, directions and the determinant
fD1x := fBx - fAx;
fD1y := fBy - fAy;
fD2x := fDx - fCx;
fD2y := fDy - fCy;
fDen := (fD1x * fD2y) - (fD1y * fD2x);     // 行列式 / the determinant
IF (fDen <> fDen) OR (ABS(fDen) > DL_FIN_LIM) THEN
    bError := TRUE;                 // 行列式非有限 / the determinant is not finite
    RETURN;
END_IF
IF ABS(fDen) < DL_EPS THEN
    bError := TRUE;                 // 平行或重合，交点不唯一 / parallel or coincident, no unique point
    RETURN;
END_IF

// 段 4｜解参数 t、u：分母已在段 3 证为非零 / segment 4, solve the two parameters
fT := (((fCx - fAx) * fD2y) - ((fCy - fAy) * fD2x)) / fDen;   // 线段一参数 / parameter on the first segment
fU := (((fCx - fAx) * fD1y) - ((fCy - fAy) * fD1x)) / fDen;   // 线段二参数 / parameter on the second segment

// 段 5｜线段域闸：任一参数越出 [0,1] 即延长线相交，按正常无交点处置 / segment 5, the segment domain gate
IF (fT < -DL_EPS) OR (fT > (DL_ONE + DL_EPS)) OR (fU < -DL_EPS) OR (fU > (DL_ONE + DL_EPS)) THEN
    RETURN;                         // bError 保持 FALSE，属正常无交点 / bError stays FALSE, this is a normal miss
END_IF

// 段 6｜交点与出口 / segment 6, the intersection point and the exit
fX := fAx + (fT * fD1x);            // 交点 X / intersection X
fY := fAy + (fT * fD1y);            // 交点 Y / intersection Y
bValid := TRUE;                     // 交点可用 / the point is usable
FC_DL_GeoLineIntersectXY := TRUE;   // 线段真实相交 / the segments really intersect
END_FUNCTION

(* ---- FC_DL_IntDivModSafe.st ---- *)
(*==============================================================================
 * 组件名称 : FC_DL_IntDivModSafe ｜ 子库 : DL_MathData ｜ v1.0.0 ｜ 2026-11-24
 * 平台     : CODESYS 3.5 / TwinCAT 3 / InoProShop / Machine Expert（纯 IEC，无厂商库）
 * 功能简介 : 有符号整数安全除余。一次算出商与余，两个出口同时给出，供定点换算、
 *            分段取模、脉冲计数分配使用。余数按「被除数符号」口径：nRem = 被除数 − 商 × 除数。
 * 契约     : 合法时返回 TRUE；nDen = 0 返回 FALSE、bError := TRUE、两出参置 0；
 *            nNum = DINT 下界且 nDen = −1 时商不可表示（−(−2^31) 回绕），
 *            返回 FALSE、bError := TRUE、两出参置 0。
 * 依赖     : 无 DL_ 内部依赖（R16 自足实现），无标准库函数调用
 * 错误码   : R297 零码位范式：eErr 恒 0，仅以 bError / bValid 表达
 * 红线自检 : R1 零全局 R2 零%I/%Q R3 纯IEC R4 除零前置 + 下界除 −1 溢出特判
 *            R5 双语注释 R6 N/A（无状态机）R7 N/A（无定时器/沿实例）
 *            R10 无类型转换 R11 全声明行分号 R15 标识符零保留字冲突 R18 N/A（无 bReset）
 * 遗留假设 : 商向零截断（IEC 61131-3 整数除法语义），余数与被除数同号；
 *            负数取余口径在不同平台有二分争议，本件以「被除数 − 商 × 除数」自证，不依赖平台取余。
 * 修订历史 : 2026-11-24 R79-A 首版（整数数论族 6/8）
 *============================================================================*)
FUNCTION FC_DL_IntDivModSafe : BOOL
VAR_INPUT
    nNum        : DINT;     // 被除数，全域 [无量纲] / dividend over the whole signed range
    nDen        : DINT;     // 除数，非零 [无量纲] / divisor, must be non zero
END_VAR
VAR_OUTPUT
    eErr        : UDINT;    // 错误码，零码位范式恒 0 / error id, always zero under the zero-code rule
    bError      : BOOL;     // 除零或商溢出为真 / TRUE on division by zero or an unrepresentable quotient
    bValid      : BOOL;     // 出参可用标志 / TRUE when the outputs are usable
    nQuot       : DINT;     // 商，向零截断，故障时 0 / quotient truncated toward zero, zero on fault
    nRem        : DINT;     // 余数，与被除数同号，故障时 0 / remainder carrying the dividend sign, zero on fault
END_VAR
VAR CONSTANT
    DL_DINT_MIN : DINT := -2147483648;  // DINT 下界，取负会回绕 [无量纲] / signed lower bound whose negation wraps
    DL_NEG_ONE  : DINT := -1;           // 负一，下界除它商不可表示 / minus one, the quotient of the lower bound overflows
    DL_ZERO     : DINT := 0;            // 整数零哨兵 / integer zero sentinel
END_VAR
VAR
    nQ          : DINT;     // 商中间量 / quotient interim value
END_VAR

// 段 1｜出口预置 / segment 1, preset the exit
FC_DL_IntDivModSafe := FALSE;   // 缺省失败 / default failure
eErr    := 0;                   // 零码位范式 / zero-code rule
bError  := FALSE;               // 预置无故障 / preset no fault
bValid  := FALSE;               // 域闸前不认出参 / the outputs are unusable until the gates pass
nQuot   := DL_ZERO;             // 商清零 / clear the quotient
nRem    := DL_ZERO;             // 余数清零 / clear the remainder

// 段 2｜除零域闸：除法前唯一必需的拦截 / segment 2, the division by zero gate
IF nDen = DL_ZERO THEN
    bError := TRUE;             // 除零 / division by zero
    RETURN;                     // 出参保持 0 / the outputs stay zero
END_IF

// 段 3｜溢出特判：下界除 −1 的商为 2^31，超出 DINT 正向上界 / segment 3, the unrepresentable quotient
IF (nNum = DL_DINT_MIN) AND (nDen = DL_NEG_ONE) THEN
    bError := TRUE;             // 商不可表示 / the quotient cannot be represented
    RETURN;                     // 出参保持 0 / the outputs stay zero
END_IF

// 段 4｜商与余：余数由乘法反算自证，不依赖平台负数取余口径 / segment 4, the quotient and a self proven remainder
nQ    := nNum / nDen;           // 商，向零截断 / quotient truncated toward zero
nQuot := nQ;                    // 出口 / publish the quotient
nRem  := nNum - (nQ * nDen);    // 余数 = 被除数 − 商 × 除数 / remainder from the product reflection
bValid := TRUE;                 // 出参可用 / the outputs are usable
FC_DL_IntDivModSafe := TRUE;    // 除余完成 / the division completed
END_FUNCTION

(* ---- FC_DL_IntSignExtractLreal.st ---- *)
(*==============================================================================
 * 组件名称 : FC_DL_IntSignExtractLreal ｜ 子库 : DL_MathData ｜ v1.0.0 ｜ 2026-11-24
 * 平台     : CODESYS 3.5 / TwinCAT 3 / InoProShop / Machine Expert（纯 IEC，无厂商库）
 * 功能简介 : 实数符号提取 —— 返回 −1 / 0 / +1 三值符号。零死区 1.0E-12 内的输入统一归 0，
 *            避免控制量在零附近因浮点噪声来回翻符号（阀门抖动、积分反向积分）。
 * 契约     : 返回 −1 / 0 / +1；非有限值（NaN 或 |x| > 1.0E308）返回 0、bError := TRUE、
 *            bValid := FALSE。纯函数无状态。
 * 依赖     : 无 DL_ 内部依赖（R16 自足实现）；Standard.library: ABS
 * 错误码   : R297 零码位范式：eErr 恒 0，仅以 bError / bValid 表达
 * 红线自检 : R1 零全局 R2 零%I/%Q R3 纯IEC R4 NaN 用自反判据 x<>x、无穷用 1.0E308 上界、
 *            零死区常量化、浮点无等号判等 R5 双语注释 R6 N/A（无状态机）
 *            R7 N/A（无定时器/沿实例）R10 无类型转换 R11 全声明行分号
 *            R15 标识符零保留字冲突 R18 N/A（无 bReset）
 * 遗留假设 : 无穷判据取 |x| > 1.0E308（LREAL 最大有限值约 1.8E308），
 *            与「用 x−x 自判」的写法互斥 —— 后者在优化编译下可能被常量折叠，已被 R77 列为死谓词。
 * 修订历史 : 2026-11-24 R79-A 首版（整数数论族 7/8）
 *============================================================================*)
FUNCTION FC_DL_IntSignExtractLreal : DINT
VAR_INPUT
    fVal        : LREAL;    // 待取符号的实数 [工程单位] / value whose sign is requested [engineering unit]
END_VAR
VAR_OUTPUT
    eErr        : UDINT;    // 错误码，零码位范式恒 0 / error id, always zero under the zero-code rule
    bError      : BOOL;     // 输入为非有限值时为真 / TRUE when the input is not finite
    bValid      : BOOL;     // 符号结论可用标志 / TRUE when the sign verdict is usable
END_VAR
VAR CONSTANT
    DL_EPS      : LREAL := 1.0E-12;      // 零死区容差，本件专用（比族内 1.0E-9 更紧）[工程单位] / zero deadband, tighter than the family default
    DL_FIN_LIM  : LREAL := 1.0E308;      // 有限性上界，超过按无穷处置 [工程单位] / finiteness ceiling, beyond it the value counts as infinity
    DL_ZERO     : DINT := 0;             // 符号零值 [无量纲] / the zero sign, dimensionless
    DL_POS_ONE  : DINT := 1;             // 正号值 [无量纲] / the positive sign, dimensionless
    DL_NEG_ONE  : DINT := -1;            // 负号值 [无量纲] / the negative sign, dimensionless
    DL_ZERO_L   : LREAL := 0.0;          // 实数零，仅用于严格不等比较 [工程单位] / real zero used by strict inequalities only
END_VAR
VAR
    fAbs        : LREAL;    // 输入的绝对值，供死区与有限性判定 / absolute value used by the deadband and the finiteness tests
END_VAR

// 段 1｜出口预置 / segment 1, preset the exit
FC_DL_IntSignExtractLreal := DL_ZERO;   // 缺省符号 0 / default sign zero
eErr   := 0;                            // 零码位范式 / zero-code rule
bError := FALSE;                        // 预置无故障 / preset no fault
bValid := TRUE;                         // 有限输入下结论恒可用 / the verdict is usable for every finite input

// 段 2｜NaN 自反判据：x <> x 成立即为 NaN，回绕 0 / segment 2, the self reflective NaN test
IF fVal <> fVal THEN
    bError := TRUE;                     // 非数 / not a number
    bValid := FALSE;                    // 符号结论不可用 / the sign verdict is unusable
    RETURN;
END_IF

// 段 3｜无穷判据：绝对值超有限上界即按非有限处置 / segment 3, the infinity test on the magnitude
fAbs := ABS(fVal);                      // 幅度 / magnitude
IF fAbs > DL_FIN_LIM THEN
    bError := TRUE;                     // 无穷 / infinity
    bValid := FALSE;                    // 符号结论不可用 / the sign verdict is unusable
    RETURN;
END_IF

// 段 4｜零死区：幅度不足容差即归 0，抑制零附近符号抖动 / segment 4, the zero deadband
IF fAbs < DL_EPS THEN
    RETURN;                            // 返回 0 / return zero
END_IF

// 段 5｜符号：死区外按严格不等比较，不使用等号 / segment 5, the sign outside the deadband
IF fVal > DL_ZERO_L THEN
    FC_DL_IntSignExtractLreal := DL_POS_ONE;    // 正号 / positive sign
ELSE
    FC_DL_IntSignExtractLreal := DL_NEG_ONE;    // 负号 / negative sign
END_IF
END_FUNCTION

(* ---- FC_DL_StatsMadFixed.st ---- *)
(*==============================================================================
 * 组件名称 : FC_DL_StatsMadFixed ｜ 子库 : DL_MathData ｜ v1.0.0 ｜ 2026-11-24
 * 平台     : CODESYS 3.5 / TwinCAT 3 / InoProShop / Machine Expert（纯 IEC，无厂商库）
 * 功能简介 : 定长样本的中位数绝对偏差 MAD = median(|xi − median(x)|)。
 *            MAD 对离群点不敏感，是比标准差更稳的离散度量 —— 传感器毛刺、
 *            单点跳变不会把 MAD 拉偏，适合做在线异常判据。排序用自实现插入排序，
 *            不调用未经验证的排序件（R16）。
 * 契约     : 返回 MAD（≥ 0）；nCnt < 1 时返回 0 且 bError := TRUE；nCnt > 10 钳到 10。
 *            偶数样本的中位数取中间两值的算术平均。数组定长 ARRAY[1..10]（R17）。
 * 依赖     : 无 DL_ 内部依赖（R16 自足实现）；Standard.library: ABS
 * 错误码   : R297 零码位范式：eErr 恒 0，仅以 bError / bValid 表达
 * 红线自检 : R1 零全局 R2 零%I/%Q R3 纯IEC R4 点数先钳位、局部数组下标恒在 1..10、
 *            偶数中位数除数为常量 2 ｜ R5 双语注释 R6 N/A（无状态机）
 *            R7 N/A（无定时器/沿实例）R10 无类型转换 R11 全声明行分号
 *            R15 标识符零保留字冲突 R17 定长数组 R18 N/A（无 bReset）
 * 遗留假设 : 非有限样本不剔除（MAD 的稳健性以有限样本为前提）；含 NaN 时比较全为假，
 *            排序不崩但 MAD 结果无意义 —— 调用方须先做非有限过滤。
 * 修订历史 : 2026-11-24 R79-A 首版（统计扩展族 3/8）
 *============================================================================*)
FUNCTION FC_DL_StatsMadFixed : LREAL
VAR_INPUT
    aVals   : ARRAY[1..10] OF LREAL;    // 样本数组，1..10 定长 [工程单位] / sample array of fixed length [engineering unit]
    nCnt    : INT;                      // 有效样本数，1~10，越界钳位 [个] / effective sample count from one to ten, clamped [count]
END_VAR
VAR_OUTPUT
    eErr    : UDINT;                    // 错误码，零码位范式恒 0 / error id, always zero under the zero-code rule
    bError  : BOOL;                     // 有效样本数为零为真 / TRUE when no usable sample exists
    bValid  : BOOL;                     // 结果可用标志 / result usable flag
END_VAR
VAR CONSTANT
    DL_PTS_MAX : INT := 10;             // 样本定长上限 [个] / fixed sample capacity [count]
    DL_PTS_MIN : INT := 1;              // 最少样本数 [个] / minimum sample count [count]
    DL_ONE     : INT := 1;              // 数组首下标 [个] / first array index [count]
    DL_TWO     : INT := 2;              // 偶数中位数的除数 [个] / divisor of the even median [count]
    DL_TWO_L   : LREAL := 2.0;          // 实数二，偶数中位数平均用 [无量纲] / real two used by the even median
    DL_ZERO_L  : LREAL := 0.0;          // 实数零哨兵 [工程单位] / real zero sentinel [engineering unit]
END_VAR
VAR
    aBuf    : ARRAY[1..10] OF LREAL;    // 排序用样本副本 [工程单位] / sorted copy of the samples [engineering unit]
    aDev    : ARRAY[1..10] OF LREAL;    // 绝对偏差数组 [工程单位] / absolute deviation array [engineering unit]
    nUse    : INT;                      // 钳位后的有效点数 [个] / effective point count after clamping [count]
    nMid    : INT;                      // 中位位置 [个] / the middle position [count]
    i       : INT;                      // 外层游标 [个] / outer cursor [count]
    j       : INT;                      // 内层游标 [个] / inner cursor [count]
    fKey    : LREAL;                    // 插入排序的待插值 [工程单位] / key of the insertion sort [engineering unit]
    fMed    : LREAL;                    // 样本中位数 [工程单位] / median of the samples [engineering unit]
END_VAR

// 段 1｜出口预置 / segment 1, preset the exit
FC_DL_StatsMadFixed := DL_ZERO_L;       // 缺省 0 / default zero
eErr   := 0;                            // 零码位范式 / zero-code rule
bError := FALSE;                        // 预置无故障 / preset no fault
bValid := FALSE;                        // 计算完成前不认结果 / unusable until the median walk ends

// 段 2｜点数钳位：上越界静默钳位，零样本按故障退出 / segment 2, clamp the count
nUse := nCnt;
IF nUse > DL_PTS_MAX THEN
    nUse := DL_PTS_MAX;
END_IF
IF nUse < DL_PTS_MIN THEN
    bError := TRUE;                     // 无样本可统计 / no sample to scan
    RETURN;
END_IF

// 段 3｜拷贝并插入排序：小规模（≤10）下插入排序最稳，无递归无额外内存 / segment 3, copy and insertion sort
FOR i := DL_ONE TO nUse DO
    aBuf[i] := aVals[i];                // 拷贝，保持入参只读 / copy so the input stays read only
END_FOR
FOR i := DL_TWO TO nUse DO
    fKey := aBuf[i];                    // 待插值 / the key to insert
    j    := i - DL_ONE;
    WHILE (j >= DL_ONE) AND (aBuf[j] > fKey) DO
        aBuf[j + DL_ONE] := aBuf[j];    // 后移空位 / shift right to open a slot
        j := j - DL_ONE;
    END_WHILE
    aBuf[j + DL_ONE] := fKey;           // 落位 / drop the key in place
END_FOR

// 段 4｜样本中位数：奇数取正中，偶数取中间两值平均 / segment 4, the median of the samples
IF (nUse MOD DL_TWO) = DL_ONE THEN
    nMid := (nUse + DL_ONE) / DL_TWO;                   // 正中位置 / the exact middle
    fMed := aBuf[nMid];
ELSE
    nMid := nUse / DL_TWO;                              // 中间左侧位置 / the left middle
    fMed := (aBuf[nMid] + aBuf[nMid + DL_ONE]) / DL_TWO_L;
END_IF

// 段 5｜绝对偏差数组：|xi − 中位数| / segment 5, the absolute deviation array
FOR i := DL_ONE TO nUse DO
    aDev[i] := ABS(aBuf[i] - fMed);
END_FOR

// 段 6｜偏差再排序，其中位数即 MAD / segment 6, sort the deviations and take their median
FOR i := DL_TWO TO nUse DO
    fKey := aDev[i];
    j    := i - DL_ONE;
    WHILE (j >= DL_ONE) AND (aDev[j] > fKey) DO
        aDev[j + DL_ONE] := aDev[j];
        j := j - DL_ONE;
    END_WHILE
    aDev[j + DL_ONE] := fKey;
END_FOR
IF (nUse MOD DL_TWO) = DL_ONE THEN
    nMid := (nUse + DL_ONE) / DL_TWO;
    FC_DL_StatsMadFixed := aDev[nMid];                  // 奇数取正中 / odd counts take the exact middle
ELSE
    nMid := nUse / DL_TWO;
    FC_DL_StatsMadFixed := (aDev[nMid] + aDev[nMid + DL_ONE]) / DL_TWO_L;   // 偶数取中间两值平均 / even counts average the middle pair
END_IF
bValid := TRUE;                                         // 结果可用 / the result is usable
END_FUNCTION

(* ---- FC_DL_StatsTrimmedMeanFixed.st ---- *)
(*==============================================================================
 * 组件名称 : FC_DL_StatsTrimmedMeanFixed ｜ 子库 : DL_MathData ｜ v1.0.0 ｜ 2026-11-24
 * 平台     : CODESYS 3.5 / TwinCAT 3 / InoProShop / Machine Expert（纯 IEC，无厂商库）
 * 功能简介 : 定长样本的截尾均值（trimmed mean）—— 先排序，两侧各去掉 nTrimEachSide 个
 *            极值，再对剩余求算术平均。截尾均值同时抗离群点与保留分布信息，
 *            是比全样本均值更稳的过程中心估计，常用于称重剔除工位与温度场均衡判定。
 * 契约     : 返回截尾均值；nCnt < 1 时返回 0 且 bError := TRUE；nCnt > 10 钳到 10；
 *            nTrimEachSide 自动钳到 0~(nCnt−1)/2，保证至少留 1 个样本参与平均。
 *            排序用自实现插入排序，数组定长 ARRAY[1..10]（R17）。
 * 依赖     : 无 DL_ 内部依赖（R16 自足实现），无标准库函数调用
 * 错误码   : R297 零码位范式：eErr 恒 0，仅以 bError / bValid 表达
 * 红线自检 : R1 零全局 R2 零%I/%Q R3 纯IEC R4 点数与截尾数双钳位、剩余样本数恒 ≥ 1 后
 *            才做除法 ｜ R5 双语注释 R6 N/A（无状态机）R7 N/A（无定时器/沿实例）
 *            R10 无类型转换 R11 全声明行分号 R15 标识符零保留字冲突
 *            R17 定长数组 R18 N/A（无 bReset）
 * 修订历史 : 2026-11-24 R79-A 首版（统计扩展族 4/8）
 *============================================================================*)
FUNCTION FC_DL_StatsTrimmedMeanFixed : LREAL
VAR_INPUT
    aVals    : ARRAY[1..10] OF LREAL;   // 样本数组，1..10 定长 [工程单位] / sample array of fixed length [engineering unit]
    nCnt     : INT;                     // 有效样本数，1~10，越界钳位 [个] / effective sample count from one to ten, clamped [count]
    nTrimEachSide : INT;                // 每侧截去的极值个数，自动钳位 [个] / values trimmed from each side, clamped [count]
END_VAR
VAR_OUTPUT
    eErr     : UDINT;                   // 错误码，零码位范式恒 0 / error id, always zero under the zero-code rule
    bError   : BOOL;                    // 有效样本数为零为真 / TRUE when no usable sample exists
    bValid   : BOOL;                    // 结果可用标志 / result usable flag
END_VAR
VAR CONSTANT
    DL_PTS_MAX : INT := 10;             // 样本定长上限 [个] / fixed sample capacity [count]
    DL_PTS_MIN : INT := 1;              // 最少样本数 [个] / minimum sample count [count]
    DL_ONE     : INT := 1;              // 数组首下标 [个] / first array index [count]
    DL_TWO     : INT := 2;              // 截尾上限式的除数 [个] / divisor of the trim cap [count]
    DL_ZERO    : INT := 0;              // 整数零哨兵 / integer zero sentinel
    DL_ZERO_L  : LREAL := 0.0;          // 实数零哨兵 [工程单位] / real zero sentinel [engineering unit]
END_VAR
VAR
    aBuf     : ARRAY[1..10] OF LREAL;   // 排序后的样本副本 [工程单位] / sorted copy of the samples [engineering unit]
    nUse     : INT;                     // 钳位后的有效点数 [个] / effective point count after clamping [count]
    nTrim    : INT;                     // 钳位后的单侧截尾数 [个] / effective trim per side [count]
    nKeep    : INT;                     // 截尾后剩余样本数 [个] / samples left after trimming [count]
    i        : INT;                     // 外层游标 [个] / outer cursor [count]
    j        : INT;                     // 内层游标 [个] / inner cursor [count]
    fKey     : LREAL;                   // 插入排序待插值 [工程单位] / key of the insertion sort [engineering unit]
    fSum     : LREAL;                   // 剩余样本累加 [工程单位] / accumulated sum of the kept samples [engineering unit]
END_VAR

// 段 1｜出口预置 / segment 1, preset the exit
FC_DL_StatsTrimmedMeanFixed := DL_ZERO_L;   // 缺省 0 / default zero
eErr   := 0;                                // 零码位范式 / zero-code rule
bError := FALSE;                            // 预置无故障 / preset no fault
bValid := FALSE;                            // 计算完成前不认结果 / unusable until the average ends

// 段 2｜点数钳位：上越界静默钳位，零样本按故障退出 / segment 2, clamp the count
nUse := nCnt;
IF nUse > DL_PTS_MAX THEN
    nUse := DL_PTS_MAX;
END_IF
IF nUse < DL_PTS_MIN THEN
    bError := TRUE;                         // 无样本可统计 / no sample to scan
    RETURN;
END_IF

// 段 3｜截尾数钳位：单侧最多去到只剩 1 个样本 / segment 3, clamp the trim so that one sample survives
nTrim := nTrimEachSide;
IF nTrim < DL_ZERO THEN
    nTrim := DL_ZERO;                       // 负截尾按 0 处理 / a negative trim means none
END_IF
IF nTrim > ((nUse - DL_ONE) / DL_TWO) THEN
    nTrim := (nUse - DL_ONE) / DL_TWO;      // 单侧上限，保证剩余至少 1 个 / the cap that keeps one sample alive
END_IF
nKeep := nUse - (DL_TWO * nTrim);           // 剩余样本数，恒 ≥ 1 / the kept count, always at least one

// 段 4｜拷贝并插入排序：升序，极值集中在两端以便截尾 / segment 4, copy and insertion sort in ascending order
FOR i := DL_ONE TO nUse DO
    aBuf[i] := aVals[i];                    // 拷贝，保持入参只读 / copy so the input stays read only
END_FOR
FOR i := DL_TWO TO nUse DO
    fKey := aBuf[i];
    j    := i - DL_ONE;
    WHILE (j >= DL_ONE) AND (aBuf[j] > fKey) DO
        aBuf[j + DL_ONE] := aBuf[j];        // 后移空位 / shift right to open a slot
        j := j - DL_ONE;
    END_WHILE
    aBuf[j + DL_ONE] := fKey;               // 落位 / drop the key in place
END_FOR

// 段 5｜截尾求和：下标 (1+nTrim) ~ (nUse−nTrim)，不会越界 / segment 5, sum the kept window
fSum := DL_ZERO_L;
FOR i := (DL_ONE + nTrim) TO (nUse - nTrim) DO
    fSum := fSum + aBuf[i];
END_FOR

// 段 6｜出口：剩余数已证 ≥ 1，除法安全 / segment 6, the divisor is proven to be at least one
FC_DL_StatsTrimmedMeanFixed := fSum / INT_TO_LREAL(nKeep);   // 截尾均值 / the trimmed mean
bValid := TRUE;                                              // 结果可用 / the result is usable
END_FUNCTION

(* ---- FB_DL_StatsSkewKurtStream.st ---- *)
(*==============================================================================
 * 组件名称 : FB_DL_StatsSkewKurtStream ｜ 子库 : DL_MathData ｜ v1.0.0 ｜ 2026-11-24
 * 平台     : CODESYS 3.5 / TwinCAT 3 / InoProShop / Machine Expert（纯 IEC，无厂商库）
 * 功能简介 : 流式三阶/四阶中心矩累加器（Terriberry 单遍递推），出偏度与超额峰度。
 *            在 Welford 的 n / mean / M2 之上再加 M3 / M4，四个量同拍更新：
 *            d = x − mean；dn = d/n；t1 = d·dn·(n−1)；
 *            M4 += t1·dn²·(n²−3n+3) + 6·dn²·M2 − 4·dn·M3；
 *            M3 += t1·dn·(n−2) − 3·dn·M2；M2 += t1；mean += dn。
 *            更新顺序固定为 M4 → M3 → M2，保证每一步读到的都是上一拍的历史矩。
 * 契约     : 偏度 = √n·M3 / M2^1.5；超额峰度 = n·M4 / M2² − 3。
 *            n < 4 时 fSkew / fKurt 置 0 且 bValid := FALSE（四阶矩少于四样本无意义）；
 *            M2 < 1.0E-18（零方差流）时形状量置 0，除零结构性不可达。
 *            bEnable 上升沿采样一次，bReset 上升沿全清（R18 / R7 均用 R_TRIG）。
 * 依赖     : 无 DL_ 内部依赖（R16 自足实现）；Standard.library: R_TRIG / ABS / SQRT
 * 错误码   : R297 零码位范式：eErr 恒 0，丢弃以 bRejected 表达
 * 红线自检 : R1 零全局 R2 零%I/%Q R3 纯IEC R4 除零前置（n≥1、M2 阈值闸）、NaN 自反判据、
 *            无穷上界、平方项先转实数再乘 ｜ R5 双语注释 R6 ENUM+CASE+ELSE 兜底
 *            R7 R_TRIG 置于 CASE 外无条件刷新 ｜ R10 标准转换 R11 全声明行分号
 *            R14 无 PROPERTY R15 标识符零保留字冲突 R18 bReset 走 R_TRIG
 * 修订历史 : 2026-11-24 R79-A 首版（统计扩展族 2/8）
 *============================================================================*)
TYPE E_DL_SkewKurtStage :
(
    eSkewIdle  := 0,        // 零样本 / no sample
    eSkewAccum := 1,        // 一至三样本，形状量不可用 / one to three samples, the shape measures are unavailable
    eSkewReady := 2         // 四样本以上，偏度峰度可用 / four samples or more, skewness and kurtosis are usable
);
END_TYPE

FUNCTION_BLOCK FB_DL_StatsSkewKurtStream
VAR_INPUT
    bEnable   : BOOL;   // 采样使能，上升沿表示新样本到达 / capture enable, a rising edge marks a new sample
    bReset    : BOOL;   // 复位，上升沿清零四个矩累加器 / reset, a rising edge clears all four moments
    fSample   : LREAL;  // 样本值，非有限者被丢弃 [工程单位] / sample value, non finite ones are dropped [engineering unit]
END_VAR
VAR_OUTPUT
    eErr      : UDINT;  // 错误码，零码位范式恒 0 / error id, always zero under the zero-code rule
    bError    : BOOL;   // 故障标志，本件不产生故障级 / fault flag, never raised by this component
    bRejected : BOOL;   // 本拍样本被丢弃（非有限） / TRUE when this cycle sample was dropped
    fMean     : LREAL;  // 在线均值 [工程单位] / running mean [engineering unit]
    fSkew     : LREAL;  // 偏度（三阶标准化矩） [无量纲] / skewness, the standardised third moment [dimensionless]
    fKurt     : LREAL;  // 超额峰度，正态分布为 0 [无量纲] / excess kurtosis, zero for a normal distribution [dimensionless]
    nCount    : UDINT;  // 已纳入样本数 [个] / number of accepted samples [count]
    bValid    : BOOL;   // n ≥ 4 时为真 / TRUE from four samples on
    eStage    : E_DL_SkewKurtStage; // 累加器阶段 / accumulator stage
END_VAR
VAR CONSTANT
    DL_ONE      : UDINT := 1;           // 无符号一 / unsigned one
    DL_FOUR     : UDINT := 4;           // 无符号四，形状量可用门槛 [个] / unsigned four, the shape measure threshold [count]
    DL_M2_MIN   : LREAL := 1.0E-18;     // 零方差闸，低于它形状量置 0 / zero variance gate
    DL_KURT_BIAS : LREAL := 3.0;        // 峰度的正态基准值 3，超额峰度需减去 [无量纲] / normal reference of the raw kurtosis [dimensionless]
    DL_THREE    : LREAL := 3.0;         // 递推式常数 3 [无量纲] / recursion constant three [dimensionless]
    DL_FOUR_L   : LREAL := 4.0;         // 递推式常数 4 [无量纲] / recursion constant four [dimensionless]
    DL_SIX      : LREAL := 6.0;         // 递推式常数 6 [无量纲] / recursion constant six [dimensionless]
    DL_ONE_L    : LREAL := 1.0;         // 实数一，用于 n−1 / real one used by the n minus one factor
    DL_TWO_L    : LREAL := 2.0;         // 实数二，用于 n−2 / real two used by the n minus two factor
    DL_FIN_LIM  : LREAL := 1.0E308;     // 有限性上界，超过按无穷处置 [工程单位] / finiteness ceiling [engineering unit]
    DL_ZERO_L   : LREAL := 0.0;         // 实数零哨兵 / real zero sentinel
END_VAR
VAR
    rtReset   : R_TRIG; // 复位上升沿检测，无条件周期刷新 / reset rising edge, refreshed every cycle
    rtSample  : R_TRIG; // 采样上升沿检测，无条件周期刷新 / sample rising edge, refreshed every cycle
    nAcc      : UDINT;  // 内部样本计数 / internal sample counter
    fMeanInt  : LREAL;  // 内部均值累加器 [工程单位] / internal mean accumulator [engineering unit]
    fM2       : LREAL;  // 二阶中心矩 [工程单位²] / second central moment [unit squared]
    fM3       : LREAL;  // 三阶中心矩 [工程单位³] / third central moment [unit cubed]
    fM4       : LREAL;  // 四阶中心矩 [工程单位⁴] / fourth central moment [unit to the fourth]
    fDelta    : LREAL;  // 新样本偏差 d [工程单位] / deviation of the new sample [engineering unit]
    fDeltaN   : LREAL;  // 偏差除以 n [工程单位] / deviation over the sample count [engineering unit]
    fTerm1    : LREAL;  // 递推主项 t1 = d·dn·(n−1) [工程单位²] / the leading recursion term [unit squared]
    fN        : LREAL;  // 样本数的实数形式 [个] / the sample count as a real number [count]
END_VAR

// 段 1｜沿检测无条件周期刷新（R7） / segment 1, refresh both edges unconditionally
rtReset(CLK := bReset);
rtSample(CLK := bEnable);

// 段 2｜出口预置 / segment 2, preset the single cycle outputs
eErr      := 0;             // 零码位范式 / zero-code rule
bError    := FALSE;         // 本件不产生故障级 / this component raises no fault
bRejected := FALSE;         // 本拍未丢弃 / nothing dropped yet

// 段 3｜复位优先：四个矩全清 / segment 3, reset has priority and clears all four moments
IF rtReset.Q THEN
    nAcc     := 0;
    fMeanInt := DL_ZERO_L;
    fM2      := DL_ZERO_L;
    fM3      := DL_ZERO_L;
    fM4      := DL_ZERO_L;
END_IF

// 段 4｜采样与递推：顺序固定 M4 → M3 → M2，均读历史矩 / segment 4, the recursion in a fixed order
IF rtSample.Q THEN
    IF (fSample <> fSample) OR (ABS(fSample) > DL_FIN_LIM) THEN
        bRejected := TRUE;                                  // 非数或无穷，丢弃 / not a number or infinity, dropped
    ELSE
        nAcc     := nAcc + DL_ONE;                          // 先自增，保证除数 ≥ 1 / increment first so the divisor is at least one
        fN       := UDINT_TO_LREAL(nAcc);                   // 实数样本数 / the count as a real number
        fDelta   := fSample - fMeanInt;                     // 偏差 / deviation
        fDeltaN  := fDelta / fN;                            // 偏差除以 n / deviation over the count
        fTerm1   := fDelta * fDeltaN * (fN - DL_ONE_L);     // 递推主项 / the leading term
        fMeanInt := fMeanInt + fDeltaN;                     // 均值递推 / mean update
        fM4      := fM4 + (fTerm1 * fDeltaN * fDeltaN * ((fN * fN) - (DL_THREE * fN) + DL_THREE)) + (DL_SIX * fDeltaN * fDeltaN * fM2) - (DL_FOUR_L * fDeltaN * fM3);
        fM3      := fM3 + (fTerm1 * fDeltaN * (fN - DL_TWO_L)) - (DL_THREE * fDeltaN * fM2);
        fM2      := fM2 + fTerm1;                           // 二阶矩最后更新，供下一拍使用 / the second moment is updated last
    END_IF
END_IF

// 段 5｜阶段机与出口发布：每分支内自洽，无跨分支残留 / segment 5, the stage machine
CASE eStage OF
    eSkewIdle, eSkewAccum:
        fMean  := fMeanInt;                         // 空相时内部均值恒 0，两相共用一条发布路径 / the internal mean is zero when empty, so both stages share one path
        fSkew  := DL_ZERO_L;                        // 不足四样本，偏度置 0 / fewer than four samples, skewness is zero
        fKurt  := DL_ZERO_L;                        // 不足四样本，峰度置 0 / fewer than four samples, kurtosis is zero
        bValid := FALSE;                            // 形状量不可用 / the shape measures are unavailable
        IF nAcc >= DL_FOUR THEN
            eStage := eSkewReady;                   // 进入可用相 / enter the ready stage
        ELSIF nAcc = 0 THEN
            eStage := eSkewIdle;                    // 回落空闲相（复位后）/ fall back to idle after a reset
        ELSE
            eStage := eSkewAccum;                   // 停在累加相 / stay at the accumulation stage
        END_IF
    eSkewReady:
        fMean := fMeanInt;
        fN    := UDINT_TO_LREAL(nAcc);              // 实数样本数 / the count as a real number
        IF fM2 > DL_M2_MIN THEN
            fSkew := (SQRT(fN) * fM3) / (fM2 * SQRT(fM2));      // √n·M3 / M2^1.5 / the standardised third moment
            fKurt := ((fN * fM4) / (fM2 * fM2)) - DL_KURT_BIAS; // n·M4 / M2² − 3 / the excess kurtosis
        ELSE
            fSkew := DL_ZERO_L;                     // 零方差流，形状量置 0（除零不可达）/ zero variance keeps the shapes at zero
            fKurt := DL_ZERO_L;
        END_IF
        bValid := TRUE;                             // 形状量可用 / the shape measures are usable
        IF nAcc < DL_FOUR THEN
            IF nAcc = 0 THEN
                eStage := eSkewIdle;                // 复位后回落 / fall back after a reset
            ELSE
                eStage := eSkewAccum;               // 回落累加相 / fall back to the accumulation stage
            END_IF
        END_IF
ELSE
    eStage := eSkewIdle;                            // 非法阶段拦截并复位 / intercept an illegal stage and recover
    fMean  := DL_ZERO_L;
    fSkew  := DL_ZERO_L;
    fKurt  := DL_ZERO_L;
    bValid := FALSE;
END_CASE

// 段 6｜计数出口：与阶段机解耦 / segment 6, publish the count independently
nCount := nAcc;
END_FUNCTION_BLOCK
